FUNCTION_BLOCK FB_STOEBERSDS_Drive_REF
VAR_INPUT
	stTerminalState			AT %I*:ST_TerminalState;
	stStoeberToPlc			AT %I*:ST_STOEBERTOPLC;
	stPlcToStoeber			AT %Q*:ST_PLCTOSTOEBER;
END_VAR
VAR_OUTPUT

END_VAR
VAR_IN_OUT

END_VAR
VAR

END_VAR

;

END_FUNCTION_BLOCK

(* stored: Version 1.1.0.1, ProductVersion 3.1.4024.15
   POU FB_STOEBERSDS_Drive_REF: Id {be8e1d2a-8871-4ca6-9d7d-a4eb80c3883c}, SpecialFunc None *)
